TYPE ST_PolarIIChamber_ArmServiceStatus :
STRUCT
	Lift : ST_PolarIIChamber_LiftTopDownServiceStatus;
	Rotate : ST_PolarIIChamber_ArmRotateServiceStatus;
	Nozzle : ARRAY[1..3] OF ST_PolarIIChamber_NozzleSupplyServiceStatus; // Unsupported elements keep ServiceId = 0.
	NozzlePort : ST_PolarIIChamber_NozzlePortServiceStatus; // Arm3/Arm4 members keep ServiceId = 0.
END_STRUCT
END_TYPE

(* stored: Version 1.1.0.1, ProductVersion 3.1.4026.18
   DUT ST_PolarIIChamber_ArmServiceStatus: Id {14000000-0000-0000-0000-000000000060} *)
